TYPE ST_GFX4IR_REF_1 : FB_GFX4IR_REF;
END_TYPE

(* stored: Version 1.1.0.1, ProductVersion 3.1.4024.15
   DUT ST_GFX4IR_REF_1: Id {5b80a7dc-e61f-4fff-a0e6-7d8353272631} *)
